PROGRAM MAIN
VAR
    fbHouse : FB_House;
END_VAR

fbHouse();

END_PROGRAM

(* stored: Version 1.1.0.1, ProductVersion 3.1.4026.20
   POU MAIN: Id {99999999-9999-4999-8999-999999999999} *)
